TYPE ET_Gr01HomeAxis :
(
	ET_Gr01HomeAxis_eWaitExecute := 0,
	ET_Gr01HomeAxis_eWaitAxisStatus,
	ET_Gr01HomeAxis_eMoveStop,
	ET_Gr01HomeAxis_eWFMoveStop,
	ET_Gr01HomeAxis_eAxisReset,
	ET_Gr01HomeAxis_eWfAxisReset,
	ET_Gr01HomeAxis_eChkAxisCoupled,
	ET_Gr01HomeAxis_eAxisRef,
	ET_Gr01HomeAxis_eWfAxisRef,
	ET_Gr01HomeAxis_eWfErrorByReference,
	ET_Gr01HomeAxis_eAxisMoveHomePos,
	ET_Gr01HomeAxis_eAxisInHomePos,
	ET_Gr01HomeAxis_eAxisSetHome,
	ET_Gr01HomeAxis_eWfSetHome,
	ET_Gr01HomeAxis_eDone := 197,
	ET_Gr01HomeAxis_eError := 198,
	ET_Gr01HomeAxis_eNoExecute := 199
);
END_TYPE

(* stored: Version 1.1.0.1, ProductVersion 3.1.4024.15
   DUT ET_Gr01HomeAxis: Id {13368119-26cc-47df-9a54-dd5fa48bc7ea} *)
